ABB RAPID module: TgtProg.mod

%%%
  VERSION:1
  LANGUAGE:ENGLISH
%%%
MODULE MOD_TgtProg

    ! -------------------------------
    ! Define customized variables here
    ! ...

	! Tool variables:

	! Reference variables:

	PROC Main()
		ConfJ \On;
		ConfL \Off;
		! Program generated by RoboDK v6.0.7 for ABB IRB 4600-60/2.05 on XX/XX/XXXX 18:00:00
		! Using nominal kinematics.
		MoveAbsJ [[10.000000,-20.000000,30.000000,-40.000000,50.000000,-60.000000],[500.000000,9E+09,9E+09,9E+09,9E+09,9E+09]],v500,z1,tool0 \WObj:=wobj0;
		MoveL [[500.000,100.000,400.000],[0.00000000,0.00000000,1.00000000,0.00000000],[0,0,0,0],[250.000000,9E+09,9E+09,9E+09,9E+09,9E+09]],v500,z1,tool0 \WObj:=wobj0;
	ENDPROC

ENDMODULE
